Yaskawa INFORM job: VEGG1.JBI

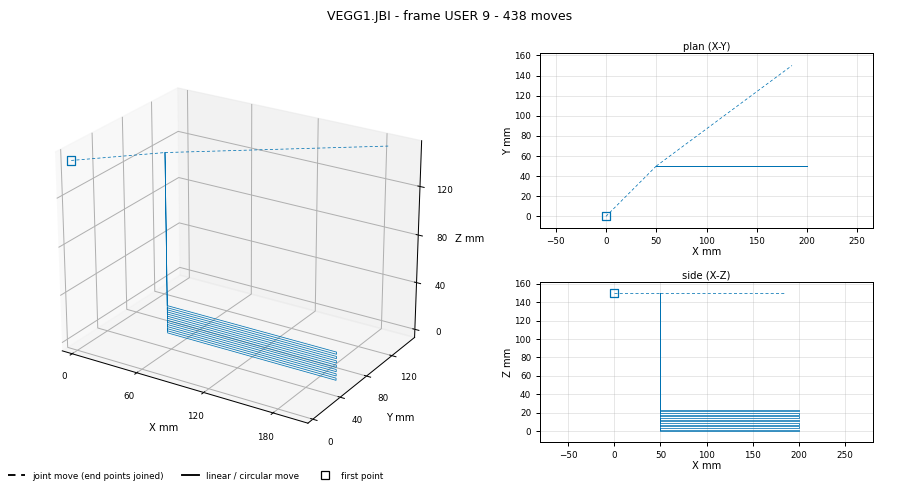
[picture p0: tool path of VEGG1.JBI in frame USER 9, 438 of 438 moves have a stored position in this frame; points joined in program order, loops and branches not executed]
/JOB
//NAME VEGG1
//POS
///NPOS 438,0,0,0,0,0
///USER 9
///TOOL 1
///POSTYPE USER
///RECTAN
///RCONF 1,0,0,0,0,0,0,0,0,0,0,0,0,0,0,0,0,0,0,0,0,0,0,0
C00000=0.000,0.000,150.000,0.0000,0.0000,180.0000
C00001=50.000,50.000,150.000,0.0000,0.0000,180.0000
C00002=50.000,50.000,0.000,0.0000,0.0000,180.0000
C00003=55.000,50.000,0.000,0.0000,0.0000,180.0000
C00004=60.000,50.000,0.000,0.0000,0.0000,180.0000
C00005=65.000,50.000,0.000,0.0000,0.0000,180.0000
C00006=70.000,50.000,0.000,0.0000,0.0000,180.0000
C00007=75.000,50.000,0.000,0.0000,0.0000,180.0000
C00008=80.000,50.000,0.000,0.0000,0.0000,180.0000
C00009=85.000,50.000,0.000,0.0000,0.0000,180.0000
C00010=90.000,50.000,0.000,0.0000,0.0000,180.0000
C00011=95.000,50.000,0.000,0.0000,0.0000,180.0000
C00012=100.000,50.000,0.000,0.0000,0.0000,180.0000
C00013=105.000,50.000,0.000,0.0000,0.0000,180.0000
C00014=110.000,50.000,0.000,0.0000,0.0000,180.0000
C00015=115.000,50.000,0.000,0.0000,0.0000,180.0000
C00016=120.000,50.000,0.000,0.0000,0.0000,180.0000
C00017=125.000,50.000,0.000,0.0000,0.0000,180.0000
C00018=130.000,50.000,0.000,0.0000,0.0000,180.0000
C00019=135.000,50.000,0.000,0.0000,0.0000,180.0000
C00020=140.000,50.000,0.000,0.0000,0.0000,180.0000
C00021=145.000,50.000,0.000,0.0000,0.0000,180.0000
C00022=150.000,50.000,0.000,0.0000,0.0000,180.0000
C00023=155.000,50.000,0.000,0.0000,0.0000,180.0000
C00024=160.000,50.000,0.000,0.0000,0.0000,180.0000
C00025=165.000,50.000,0.000,0.0000,0.0000,180.0000
C00026=170.000,50.000,0.000,0.0000,0.0000,180.0000
C00027=175.000,50.000,0.000,0.0000,0.0000,180.0000
C00028=180.000,50.000,0.000,0.0000,0.0000,180.0000
C00029=185.000,50.000,0.000,0.0000,0.0000,180.0000
C00030=190.000,50.000,0.000,0.0000,0.0000,180.0000
C00031=195.000,50.000,0.000,0.0000,0.0000,180.0000
C00032=200.000,50.000,0.000,0.0000,0.0000,180.0000
C00033=200.000,50.000,1.800,0.0000,0.0000,180.0000
C00034=195.000,50.000,1.800,0.0000,0.0000,180.0000
C00035=190.000,50.000,1.800,0.0000,0.0000,180.0000
C00036=185.000,50.000,1.800,0.0000,0.0000,180.0000
C00037=180.000,50.000,1.800,0.0000,0.0000,180.0000
C00038=175.000,50.000,1.800,0.0000,0.0000,180.0000
C00039=170.000,50.000,1.800,0.0000,0.0000,180.0000
C00040=165.000,50.000,1.800,0.0000,0.0000,180.0000
C00041=160.000,50.000,1.800,0.0000,0.0000,180.0000
C00042=155.000,50.000,1.800,0.0000,0.0000,180.0000
C00043=150.000,50.000,1.800,0.0000,0.0000,180.0000
C00044=145.000,50.000,1.800,0.0000,0.0000,180.0000
C00045=140.000,50.000,1.800,0.0000,0.0000,180.0000
C00046=135.000,50.000,1.800,0.0000,0.0000,180.0000
C00047=130.000,50.000,1.800,0.0000,0.0000,180.0000
C00048=125.000,50.000,1.800,0.0000,0.0000,180.0000
C00049=120.000,50.000,1.800,0.0000,0.0000,180.0000
C00050=115.000,50.000,1.800,0.0000,0.0000,180.0000
C00051=110.000,50.000,1.800,0.0000,0.0000,180.0000
C00052=105.000,50.000,1.800,0.0000,0.0000,180.0000
C00053=100.000,50.000,1.800,0.0000,0.0000,180.0000
C00054=95.000,50.000,1.800,0.0000,0.0000,180.0000
C00055=90.000,50.000,1.800,0.0000,0.0000,180.0000
C00056=85.000,50.000,1.800,0.0000,0.0000,180.0000
C00057=80.000,50.000,1.800,0.0000,0.0000,180.0000
C00058=75.000,50.000,1.800,0.0000,0.0000,180.0000
C00059=70.000,50.000,1.800,0.0000,0.0000,180.0000
C00060=65.000,50.000,1.800,0.0000,0.0000,180.0000
C00061=60.000,50.000,1.800,0.0000,0.0000,180.0000
C00062=55.000,50.000,1.800,0.0000,0.0000,180.0000
C00063=50.000,50.000,1.800,0.0000,0.0000,180.0000
C00064=50.000,50.000,3.600,0.0000,0.0000,180.0000
C00065=55.000,50.000,3.600,0.0000,0.0000,180.0000
C00066=60.000,50.000,3.600,0.0000,0.0000,180.0000
C00067=65.000,50.000,3.600,0.0000,0.0000,180.0000
C00068=70.000,50.000,3.600,0.0000,0.0000,180.0000
C00069=75.000,50.000,3.600,0.0000,0.0000,180.0000
C00070=80.000,50.000,3.600,0.0000,0.0000,180.0000
C00071=85.000,50.000,3.600,0.0000,0.0000,180.0000
C00072=90.000,50.000,3.600,0.0000,0.0000,180.0000
C00073=95.000,50.000,3.600,0.0000,0.0000,180.0000
C00074=100.000,50.000,3.600,0.0000,0.0000,180.0000
C00075=105.000,50.000,3.600,0.0000,0.0000,180.0000
C00076=110.000,50.000,3.600,0.0000,0.0000,180.0000
C00077=115.000,50.000,3.600,0.0000,0.0000,180.0000
C00078=120.000,50.000,3.600,0.0000,0.0000,180.0000
C00079=125.000,50.000,3.600,0.0000,0.0000,180.0000
C00080=130.000,50.000,3.600,0.0000,0.0000,180.0000
C00081=135.000,50.000,3.600,0.0000,0.0000,180.0000
C00082=140.000,50.000,3.600,0.0000,0.0000,180.0000
C00083=145.000,50.000,3.600,0.0000,0.0000,180.0000
C00084=150.000,50.000,3.600,0.0000,0.0000,180.0000
C00085=155.000,50.000,3.600,0.0000,0.0000,180.0000
C00086=160.000,50.000,3.600,0.0000,0.0000,180.0000
C00087=165.000,50.000,3.600,0.0000,0.0000,180.0000
C00088=170.000,50.000,3.600,0.0000,0.0000,180.0000
C00089=175.000,50.000,3.600,0.0000,0.0000,180.0000
C00090=180.000,50.000,3.600,0.0000,0.0000,180.0000
C00091=185.000,50.000,3.600,0.0000,0.0000,180.0000
C00092=190.000,50.000,3.600,0.0000,0.0000,180.0000
C00093=195.000,50.000,3.600,0.0000,0.0000,180.0000
C00094=200.000,50.000,3.600,0.0000,0.0000,180.0000
C00095=200.000,50.000,5.400,0.0000,0.0000,180.0000
C00096=195.000,50.000,5.400,0.0000,0.0000,180.0000
C00097=190.000,50.000,5.400,0.0000,0.0000,180.0000
C00098=185.000,50.000,5.400,0.0000,0.0000,180.0000
C00099=180.000,50.000,5.400,0.0000,0.0000,180.0000
C00100=175.000,50.000,5.400,0.0000,0.0000,180.0000
C00101=170.000,50.000,5.400,0.0000,0.0000,180.0000
C00102=165.000,50.000,5.400,0.0000,0.0000,180.0000
C00103=160.000,50.000,5.400,0.0000,0.0000,180.0000
C00104=155.000,50.000,5.400,0.0000,0.0000,180.0000
C00105=150.000,50.000,5.400,0.0000,0.0000,180.0000
C00106=145.000,50.000,5.400,0.0000,0.0000,180.0000
C00107=140.000,50.000,5.400,0.0000,0.0000,180.0000
C00108=135.000,50.000,5.400,0.0000,0.0000,180.0000
C00109=130.000,50.000,5.400,0.0000,0.0000,180.0000
C00110=125.000,50.000,5.400,0.0000,0.0000,180.0000
C00111=120.000,50.000,5.400,0.0000,0.0000,180.0000
C00112=115.000,50.000,5.400,0.0000,0.0000,180.0000
C00113=110.000,50.000,5.400,0.0000,0.0000,180.0000
C00114=105.000,50.000,5.400,0.0000,0.0000,180.0000
C00115=100.000,50.000,5.400,0.0000,0.0000,180.0000
C00116=95.000,50.000,5.400,0.0000,0.0000,180.0000
C00117=90.000,50.000,5.400,0.0000,0.0000,180.0000
C00118=85.000,50.000,5.400,0.0000,0.0000,180.0000
C00119=80.000,50.000,5.400,0.0000,0.0000,180.0000
C00120=75.000,50.000,5.400,0.0000,0.0000,180.0000
C00121=70.000,50.000,5.400,0.0000,0.0000,180.0000
C00122=65.000,50.000,5.400,0.0000,0.0000,180.0000
C00123=60.000,50.000,5.400,0.0000,0.0000,180.0000
C00124=55.000,50.000,5.400,0.0000,0.0000,180.0000
C00125=50.000,50.000,5.400,0.0000,0.0000,180.0000
C00126=50.000,50.000,7.200,0.0000,0.0000,180.0000
C00127=55.000,50.000,7.200,0.0000,0.0000,180.0000
C00128=60.000,50.000,7.200,0.0000,0.0000,180.0000
C00129=65.000,50.000,7.200,0.0000,0.0000,180.0000
C00130=70.000,50.000,7.200,0.0000,0.0000,180.0000
C00131=75.000,50.000,7.200,0.0000,0.0000,180.0000
C00132=80.000,50.000,7.200,0.0000,0.0000,180.0000
C00133=85.000,50.000,7.200,0.0000,0.0000,180.0000
C00134=90.000,50.000,7.200,0.0000,0.0000,180.0000
C00135=95.000,50.000,7.200,0.0000,0.0000,180.0000
C00136=100.000,50.000,7.200,0.0000,0.0000,180.0000
C00137=105.000,50.000,7.200,0.0000,0.0000,180.0000
C00138=110.000,50.000,7.200,0.0000,0.0000,180.0000
C00139=115.000,50.000,7.200,0.0000,0.0000,180.0000
C00140=120.000,50.000,7.200,0.0000,0.0000,180.0000
C00141=125.000,50.000,7.200,0.0000,0.0000,180.0000
C00142=130.000,50.000,7.200,0.0000,0.0000,180.0000
C00143=135.000,50.000,7.200,0.0000,0.0000,180.0000
C00144=140.000,50.000,7.200,0.0000,0.0000,180.0000
C00145=145.000,50.000,7.200,0.0000,0.0000,180.0000
C00146=150.000,50.000,7.200,0.0000,0.0000,180.0000
C00147=155.000,50.000,7.200,0.0000,0.0000,180.0000
C00148=160.000,50.000,7.200,0.0000,0.0000,180.0000
C00149=165.000,50.000,7.200,0.0000,0.0000,180.0000
C00150=170.000,50.000,7.200,0.0000,0.0000,180.0000
C00151=175.000,50.000,7.200,0.0000,0.0000,180.0000
C00152=180.000,50.000,7.200,0.0000,0.0000,180.0000
C00153=185.000,50.000,7.200,0.0000,0.0000,180.0000
C00154=190.000,50.000,7.200,0.0000,0.0000,180.0000
C00155=195.000,50.000,7.200,0.0000,0.0000,180.0000
C00156=200.000,50.000,7.200,0.0000,0.0000,180.0000
C00157=200.000,50.000,9.000,0.0000,0.0000,180.0000
C00158=195.000,50.000,9.000,0.0000,0.0000,180.0000
C00159=190.000,50.000,9.000,0.0000,0.0000,180.0000
C00160=185.000,50.000,9.000,0.0000,0.0000,180.0000
C00161=180.000,50.000,9.000,0.0000,0.0000,180.0000
C00162=175.000,50.000,9.000,0.0000,0.0000,180.0000
C00163=170.000,50.000,9.000,0.0000,0.0000,180.0000
C00164=165.000,50.000,9.000,0.0000,0.0000,180.0000
C00165=160.000,50.000,9.000,0.0000,0.0000,180.0000
C00166=155.000,50.000,9.000,0.0000,0.0000,180.0000
C00167=150.000,50.000,9.000,0.0000,0.0000,180.0000
C00168=145.000,50.000,9.000,0.0000,0.0000,180.0000
C00169=140.000,50.000,9.000,0.0000,0.0000,180.0000
C00170=135.000,50.000,9.000,0.0000,0.0000,180.0000
C00171=130.000,50.000,9.000,0.0000,0.0000,180.0000
C00172=125.000,50.000,9.000,0.0000,0.0000,180.0000
C00173=120.000,50.000,9.000,0.0000,0.0000,180.0000
C00174=115.000,50.000,9.000,0.0000,0.0000,180.0000
C00175=110.000,50.000,9.000,0.0000,0.0000,180.0000
C00176=105.000,50.000,9.000,0.0000,0.0000,180.0000
C00177=100.000,50.000,9.000,0.0000,0.0000,180.0000
C00178=95.000,50.000,9.000,0.0000,0.0000,180.0000
C00179=90.000,50.000,9.000,0.0000,0.0000,180.0000
C00180=85.000,50.000,9.000,0.0000,0.0000,180.0000
C00181=80.000,50.000,9.000,0.0000,0.0000,180.0000
C00182=75.000,50.000,9.000,0.0000,0.0000,180.0000
C00183=70.000,50.000,9.000,0.0000,0.0000,180.0000
C00184=65.000,50.000,9.000,0.0000,0.0000,180.0000
C00185=60.000,50.000,9.000,0.0000,0.0000,180.0000
C00186=55.000,50.000,9.000,0.0000,0.0000,180.0000
C00187=50.000,50.000,9.000,0.0000,0.0000,180.0000
C00188=50.000,50.000,10.800,0.0000,0.0000,180.0000
C00189=55.000,50.000,10.800,0.0000,0.0000,180.0000
C00190=60.000,50.000,10.800,0.0000,0.0000,180.0000
C00191=65.000,50.000,10.800,0.0000,0.0000,180.0000
C00192=70.000,50.000,10.800,0.0000,0.0000,180.0000
C00193=75.000,50.000,10.800,0.0000,0.0000,180.0000
C00194=80.000,50.000,10.800,0.0000,0.0000,180.0000
C00195=85.000,50.000,10.800,0.0000,0.0000,180.0000
C00196=90.000,50.000,10.800,0.0000,0.0000,180.0000
C00197=95.000,50.000,10.800,0.0000,0.0000,180.0000
C00198=100.000,50.000,10.800,0.0000,0.0000,180.0000
C00199=105.000,50.000,10.800,0.0000,0.0000,180.0000
C00200=110.000,50.000,10.800,0.0000,0.0000,180.0000
C00201=115.000,50.000,10.800,0.0000,0.0000,180.0000
C00202=120.000,50.000,10.800,0.0000,0.0000,180.0000
C00203=125.000,50.000,10.800,0.0000,0.0000,180.0000
C00204=130.000,50.000,10.800,0.0000,0.0000,180.0000
C00205=135.000,50.000,10.800,0.0000,0.0000,180.0000
C00206=140.000,50.000,10.800,0.0000,0.0000,180.0000
C00207=145.000,50.000,10.800,0.0000,0.0000,180.0000
C00208=150.000,50.000,10.800,0.0000,0.0000,180.0000
C00209=155.000,50.000,10.800,0.0000,0.0000,180.0000
C00210=160.000,50.000,10.800,0.0000,0.0000,180.0000
C00211=165.000,50.000,10.800,0.0000,0.0000,180.0000
C00212=170.000,50.000,10.800,0.0000,0.0000,180.0000
C00213=175.000,50.000,10.800,0.0000,0.0000,180.0000
C00214=180.000,50.000,10.800,0.0000,0.0000,180.0000
C00215=185.000,50.000,10.800,0.0000,0.0000,180.0000
C00216=190.000,50.000,10.800,0.0000,0.0000,180.0000
C00217=195.000,50.000,10.800,0.0000,0.0000,180.0000
C00218=200.000,50.000,10.800,0.0000,0.0000,180.0000
C00219=200.000,50.000,12.600,0.0000,0.0000,180.0000
C00220=195.000,50.000,12.600,0.0000,0.0000,180.0000
C00221=190.000,50.000,12.600,0.0000,0.0000,180.0000
C00222=185.000,50.000,12.600,0.0000,0.0000,180.0000
C00223=180.000,50.000,12.600,0.0000,0.0000,180.0000
C00224=175.000,50.000,12.600,0.0000,0.0000,180.0000
C00225=170.000,50.000,12.600,0.0000,0.0000,180.0000
C00226=165.000,50.000,12.600,0.0000,0.0000,180.0000
C00227=160.000,50.000,12.600,0.0000,0.0000,180.0000
C00228=155.000,50.000,12.600,0.0000,0.0000,180.0000
C00229=150.000,50.000,12.600,0.0000,0.0000,180.0000
C00230=145.000,50.000,12.600,0.0000,0.0000,180.0000
C00231=140.000,50.000,12.600,0.0000,0.0000,180.0000
C00232=135.000,50.000,12.600,0.0000,0.0000,180.0000
C00233=130.000,50.000,12.600,0.0000,0.0000,180.0000
C00234=125.000,50.000,12.600,0.0000,0.0000,180.0000
C00235=120.000,50.000,12.600,0.0000,0.0000,180.0000
C00236=115.000,50.000,12.600,0.0000,0.0000,180.0000
C00237=110.000,50.000,12.600,0.0000,0.0000,180.0000
C00238=105.000,50.000,12.600,0.0000,0.0000,180.0000
C00239=100.000,50.000,12.600,0.0000,0.0000,180.0000
C00240=95.000,50.000,12.600,0.0000,0.0000,180.0000
C00241=90.000,50.000,12.600,0.0000,0.0000,180.0000
C00242=85.000,50.000,12.600,0.0000,0.0000,180.0000
C00243=80.000,50.000,12.600,0.0000,0.0000,180.0000
C00244=75.000,50.000,12.600,0.0000,0.0000,180.0000
C00245=70.000,50.000,12.600,0.0000,0.0000,180.0000
C00246=65.000,50.000,12.600,0.0000,0.0000,180.0000
C00247=60.000,50.000,12.600,0.0000,0.0000,180.0000
C00248=55.000,50.000,12.600,0.0000,0.0000,180.0000
C00249=50.000,50.000,12.600,0.0000,0.0000,180.0000
C00250=50.000,50.000,14.400,0.0000,0.0000,180.0000
C00251=55.000,50.000,14.400,0.0000,0.0000,180.0000
C00252=60.000,50.000,14.400,0.0000,0.0000,180.0000
C00253=65.000,50.000,14.400,0.0000,0.0000,180.0000
C00254=70.000,50.000,14.400,0.0000,0.0000,180.0000
C00255=75.000,50.000,14.400,0.0000,0.0000,180.0000
C00256=80.000,50.000,14.400,0.0000,0.0000,180.0000
C00257=85.000,50.000,14.400,0.0000,0.0000,180.0000
C00258=90.000,50.000,14.400,0.0000,0.0000,180.0000
C00259=95.000,50.000,14.400,0.0000,0.0000,180.0000
C00260=100.000,50.000,14.400,0.0000,0.0000,180.0000
C00261=105.000,50.000,14.400,0.0000,0.0000,180.0000
C00262=110.000,50.000,14.400,0.0000,0.0000,180.0000
C00263=115.000,50.000,14.400,0.0000,0.0000,180.0000
C00264=120.000,50.000,14.400,0.0000,0.0000,180.0000
C00265=125.000,50.000,14.400,0.0000,0.0000,180.0000
C00266=130.000,50.000,14.400,0.0000,0.0000,180.0000
C00267=135.000,50.000,14.400,0.0000,0.0000,180.0000
C00268=140.000,50.000,14.400,0.0000,0.0000,180.0000
C00269=145.000,50.000,14.400,0.0000,0.0000,180.0000
C00270=150.000,50.000,14.400,0.0000,0.0000,180.0000
C00271=155.000,50.000,14.400,0.0000,0.0000,180.0000
C00272=160.000,50.000,14.400,0.0000,0.0000,180.0000
C00273=165.000,50.000,14.400,0.0000,0.0000,180.0000
C00274=170.000,50.000,14.400,0.0000,0.0000,180.0000
C00275=175.000,50.000,14.400,0.0000,0.0000,180.0000
C00276=180.000,50.000,14.400,0.0000,0.0000,180.0000
C00277=185.000,50.000,14.400,0.0000,0.0000,180.0000
C00278=190.000,50.000,14.400,0.0000,0.0000,180.0000
C00279=195.000,50.000,14.400,0.0000,0.0000,180.0000
C00280=200.000,50.000,14.400,0.0000,0.0000,180.0000
C00281=200.000,50.000,16.200,0.0000,0.0000,180.0000
C00282=195.000,50.000,16.200,0.0000,0.0000,180.0000
C00283=190.000,50.000,16.200,0.0000,0.0000,180.0000
C00284=185.000,50.000,16.200,0.0000,0.0000,180.0000
C00285=180.000,50.000,16.200,0.0000,0.0000,180.0000
C00286=175.000,50.000,16.200,0.0000,0.0000,180.0000
C00287=170.000,50.000,16.200,0.0000,0.0000,180.0000
C00288=165.000,50.000,16.200,0.0000,0.0000,180.0000
C00289=160.000,50.000,16.200,0.0000,0.0000,180.0000
C00290=155.000,50.000,16.200,0.0000,0.0000,180.0000
C00291=150.000,50.000,16.200,0.0000,0.0000,180.0000
C00292=145.000,50.000,16.200,0.0000,0.0000,180.0000
C00293=140.000,50.000,16.200,0.0000,0.0000,180.0000
C00294=135.000,50.000,16.200,0.0000,0.0000,180.0000
C00295=130.000,50.000,16.200,0.0000,0.0000,180.0000
C00296=125.000,50.000,16.200,0.0000,0.0000,180.0000
C00297=120.000,50.000,16.200,0.0000,0.0000,180.0000
C00298=115.000,50.000,16.200,0.0000,0.0000,180.0000
C00299=110.000,50.000,16.200,0.0000,0.0000,180.0000
C00300=105.000,50.000,16.200,0.0000,0.0000,180.0000
C00301=100.000,50.000,16.200,0.0000,0.0000,180.0000
C00302=95.000,50.000,16.200,0.0000,0.0000,180.0000
C00303=90.000,50.000,16.200,0.0000,0.0000,180.0000
C00304=85.000,50.000,16.200,0.0000,0.0000,180.0000
C00305=80.000,50.000,16.200,0.0000,0.0000,180.0000
C00306=75.000,50.000,16.200,0.0000,0.0000,180.0000
C00307=70.000,50.000,16.200,0.0000,0.0000,180.0000
C00308=65.000,50.000,16.200,0.0000,0.0000,180.0000
C00309=60.000,50.000,16.200,0.0000,0.0000,180.0000
C00310=55.000,50.000,16.200,0.0000,0.0000,180.0000
C00311=50.000,50.000,16.200,0.0000,0.0000,180.0000
C00312=50.000,50.000,18.000,0.0000,0.0000,180.0000
C00313=55.000,50.000,18.000,0.0000,0.0000,180.0000
C00314=60.000,50.000,18.000,0.0000,0.0000,180.0000
C00315=65.000,50.000,18.000,0.0000,0.0000,180.0000
C00316=70.000,50.000,18.000,0.0000,0.0000,180.0000
C00317=75.000,50.000,18.000,0.0000,0.0000,180.0000
C00318=80.000,50.000,18.000,0.0000,0.0000,180.0000
C00319=85.000,50.000,18.000,0.0000,0.0000,180.0000
C00320=90.000,50.000,18.000,0.0000,0.0000,180.0000
C00321=95.000,50.000,18.000,0.0000,0.0000,180.0000
C00322=100.000,50.000,18.000,0.0000,0.0000,180.0000
C00323=105.000,50.000,18.000,0.0000,0.0000,180.0000
C00324=110.000,50.000,18.000,0.0000,0.0000,180.0000
C00325=115.000,50.000,18.000,0.0000,0.0000,180.0000
C00326=120.000,50.000,18.000,0.0000,0.0000,180.0000
C00327=125.000,50.000,18.000,0.0000,0.0000,180.0000
C00328=130.000,50.000,18.000,0.0000,0.0000,180.0000
C00329=135.000,50.000,18.000,0.0000,0.0000,180.0000
C00330=140.000,50.000,18.000,0.0000,0.0000,180.0000
C00331=145.000,50.000,18.000,0.0000,0.0000,180.0000
C00332=150.000,50.000,18.000,0.0000,0.0000,180.0000
C00333=155.000,50.000,18.000,0.0000,0.0000,180.0000
C00334=160.000,50.000,18.000,0.0000,0.0000,180.0000
C00335=165.000,50.000,18.000,0.0000,0.0000,180.0000
C00336=170.000,50.000,18.000,0.0000,0.0000,180.0000
C00337=175.000,50.000,18.000,0.0000,0.0000,180.0000
C00338=180.000,50.000,18.000,0.0000,0.0000,180.0000
C00339=185.000,50.000,18.000,0.0000,0.0000,180.0000
C00340=190.000,50.000,18.000,0.0000,0.0000,180.0000
C00341=195.000,50.000,18.000,0.0000,0.0000,180.0000
C00342=200.000,50.000,18.000,0.0000,0.0000,180.0000
C00343=200.000,50.000,19.800,0.0000,0.0000,180.0000
C00344=195.000,50.000,19.800,0.0000,0.0000,180.0000
C00345=190.000,50.000,19.800,0.0000,0.0000,180.0000
C00346=185.000,50.000,19.800,0.0000,0.0000,180.0000
C00347=180.000,50.000,19.800,0.0000,0.0000,180.0000
C00348=175.000,50.000,19.800,0.0000,0.0000,180.0000
C00349=170.000,50.000,19.800,0.0000,0.0000,180.0000
C00350=165.000,50.000,19.800,0.0000,0.0000,180.0000
C00351=160.000,50.000,19.800,0.0000,0.0000,180.0000
C00352=155.000,50.000,19.800,0.0000,0.0000,180.0000
C00353=150.000,50.000,19.800,0.0000,0.0000,180.0000
C00354=145.000,50.000,19.800,0.0000,0.0000,180.0000
C00355=140.000,50.000,19.800,0.0000,0.0000,180.0000
C00356=135.000,50.000,19.800,0.0000,0.0000,180.0000
C00357=130.000,50.000,19.800,0.0000,0.0000,180.0000
C00358=125.000,50.000,19.800,0.0000,0.0000,180.0000
C00359=120.000,50.000,19.800,0.0000,0.0000,180.0000
C00360=115.000,50.000,19.800,0.0000,0.0000,180.0000
C00361=110.000,50.000,19.800,0.0000,0.0000,180.0000
C00362=105.000,50.000,19.800,0.0000,0.0000,180.0000
C00363=100.000,50.000,19.800,0.0000,0.0000,180.0000
C00364=95.000,50.000,19.800,0.0000,0.0000,180.0000
C00365=90.000,50.000,19.800,0.0000,0.0000,180.0000
C00366=85.000,50.000,19.800,0.0000,0.0000,180.0000
C00367=80.000,50.000,19.800,0.0000,0.0000,180.0000
C00368=75.000,50.000,19.800,0.0000,0.0000,180.0000
C00369=70.000,50.000,19.800,0.0000,0.0000,180.0000
C00370=65.000,50.000,19.800,0.0000,0.0000,180.0000
C00371=60.000,50.000,19.800,0.0000,0.0000,180.0000
C00372=55.000,50.000,19.800,0.0000,0.0000,180.0000
C00373=50.000,50.000,19.800,0.0000,0.0000,180.0000
C00374=50.000,50.000,21.600,0.0000,0.0000,180.0000
C00375=55.000,50.000,21.600,0.0000,0.0000,180.0000
C00376=60.000,50.000,21.600,0.0000,0.0000,180.0000
C00377=65.000,50.000,21.600,0.0000,0.0000,180.0000
C00378=70.000,50.000,21.600,0.0000,0.0000,180.0000
C00379=75.000,50.000,21.600,0.0000,0.0000,180.0000
C00380=80.000,50.000,21.600,0.0000,0.0000,180.0000
C00381=85.000,50.000,21.600,0.0000,0.0000,180.0000
C00382=90.000,50.000,21.600,0.0000,0.0000,180.0000
C00383=95.000,50.000,21.600,0.0000,0.0000,180.0000
C00384=100.000,50.000,21.600,0.0000,0.0000,180.0000
C00385=105.000,50.000,21.600,0.0000,0.0000,180.0000
C00386=110.000,50.000,21.600,0.0000,0.0000,180.0000
C00387=115.000,50.000,21.600,0.0000,0.0000,180.0000
C00388=120.000,50.000,21.600,0.0000,0.0000,180.0000
C00389=125.000,50.000,21.600,0.0000,0.0000,180.0000
C00390=130.000,50.000,21.600,0.0000,0.0000,180.0000
C00391=135.000,50.000,21.600,0.0000,0.0000,180.0000
C00392=140.000,50.000,21.600,0.0000,0.0000,180.0000
C00393=145.000,50.000,21.600,0.0000,0.0000,180.0000
C00394=150.000,50.000,21.600,0.0000,0.0000,180.0000
C00395=155.000,50.000,21.600,0.0000,0.0000,180.0000
C00396=160.000,50.000,21.600,0.0000,0.0000,180.0000
C00397=165.000,50.000,21.600,0.0000,0.0000,180.0000
C00398=170.000,50.000,21.600,0.0000,0.0000,180.0000
C00399=175.000,50.000,21.600,0.0000,0.0000,180.0000
C00400=180.000,50.000,21.600,0.0000,0.0000,180.0000
C00401=185.000,50.000,21.600,0.0000,0.0000,180.0000
C00402=190.000,50.000,21.600,0.0000,0.0000,180.0000
C00403=195.000,50.000,21.600,0.0000,0.0000,180.0000
C00404=200.000,50.000,21.600,0.0000,0.0000,180.0000
C00405=200.000,50.000,23.400,0.0000,0.0000,180.0000
C00406=195.000,50.000,23.400,0.0000,0.0000,180.0000
C00407=190.000,50.000,23.400,0.0000,0.0000,180.0000
C00408=185.000,50.000,23.400,0.0000,0.0000,180.0000
C00409=180.000,50.000,23.400,0.0000,0.0000,180.0000
C00410=175.000,50.000,23.400,0.0000,0.0000,180.0000
C00411=170.000,50.000,23.400,0.0000,0.0000,180.0000
C00412=165.000,50.000,23.400,0.0000,0.0000,180.0000
C00413=160.000,50.000,23.400,0.0000,0.0000,180.0000
C00414=155.000,50.000,23.400,0.0000,0.0000,180.0000
C00415=150.000,50.000,23.400,0.0000,0.0000,180.0000
C00416=145.000,50.000,23.400,0.0000,0.0000,180.0000
C00417=140.000,50.000,23.400,0.0000,0.0000,180.0000
C00418=135.000,50.000,23.400,0.0000,0.0000,180.0000
C00419=130.000,50.000,23.400,0.0000,0.0000,180.0000
C00420=125.000,50.000,23.400,0.0000,0.0000,180.0000
C00421=120.000,50.000,23.400,0.0000,0.0000,180.0000
C00422=115.000,50.000,23.400,0.0000,0.0000,180.0000
C00423=110.000,50.000,23.400,0.0000,0.0000,180.0000
C00424=105.000,50.000,23.400,0.0000,0.0000,180.0000
C00425=100.000,50.000,23.400,0.0000,0.0000,180.0000
C00426=95.000,50.000,23.400,0.0000,0.0000,180.0000
C00427=90.000,50.000,23.400,0.0000,0.0000,180.0000
C00428=85.000,50.000,23.400,0.0000,0.0000,180.0000
C00429=80.000,50.000,23.400,0.0000,0.0000,180.0000
C00430=75.000,50.000,23.400,0.0000,0.0000,180.0000
C00431=70.000,50.000,23.400,0.0000,0.0000,180.0000
C00432=65.000,50.000,23.400,0.0000,0.0000,180.0000
C00433=60.000,50.000,23.400,0.0000,0.0000,180.0000
C00434=55.000,50.000,23.400,0.0000,0.0000,180.0000
C00435=50.000,50.000,23.400,0.0000,0.0000,180.0000
C00436=50.000,50.000,150.000,0.0000,0.0000,180.0000
C00437=185.000,150.000,150.000,0.0000,0.0000,180.0000
//INST
///DATE 2026/10/20 11:28
///ATTR SC,RW,RJ
////FRAME USER 9
///GROUP1 RB1
NOP
MOVJ C00000 VJ=0.78
MOVJ C00001 VJ=0.78
MOVL C00002 V=11.0 ACC=20 DEC=20
MACRO1 MJ#(0) ARGF1
ARCON
MOVL C00003 V=8.0 ACC=20 DEC=20
MOVL C00004 V=8.0 ACC=20 DEC=20
MOVL C00005 V=8.0 ACC=20 DEC=20
MOVL C00006 V=8.0 ACC=20 DEC=20
MOVL C00007 V=8.0 ACC=20 DEC=20
MOVL C00008 V=8.0 ACC=20 DEC=20
MOVL C00009 V=8.0 ACC=20 DEC=20
MOVL C00010 V=8.0 ACC=20 DEC=20
MOVL C00011 V=8.0 ACC=20 DEC=20
MOVL C00012 V=8.0 ACC=20 DEC=20
MOVL C00013 V=8.0 ACC=20 DEC=20
MOVL C00014 V=8.0 ACC=20 DEC=20
MOVL C00015 V=8.0 ACC=20 DEC=20
MOVL C00016 V=8.0 ACC=20 DEC=20
MOVL C00017 V=8.0 ACC=20 DEC=20
MOVL C00018 V=8.0 ACC=20 DEC=20
MOVL C00019 V=8.0 ACC=20 DEC=20
MOVL C00020 V=8.0 ACC=20 DEC=20
MOVL C00021 V=8.0 ACC=20 DEC=20
MOVL C00022 V=8.0 ACC=20 DEC=20
MOVL C00023 V=8.0 ACC=20 DEC=20
MOVL C00024 V=8.0 ACC=20 DEC=20
MOVL C00025 V=8.0 ACC=20 DEC=20
MOVL C00026 V=8.0 ACC=20 DEC=20
MOVL C00027 V=8.0 ACC=20 DEC=20
MOVL C00028 V=8.0 ACC=20 DEC=20
MOVL C00029 V=8.0 ACC=20 DEC=20
MOVL C00030 V=8.0 ACC=20 DEC=20
MOVL C00031 V=8.0 ACC=20 DEC=20
MOVL C00032 V=8.0 ACC=20 DEC=20
ARCOF
TIMER T=60.0
MOVL C00033 V=11.0 ACC=20 DEC=20
MACRO1 MJ#(0) ARGF2
ARCON
MOVL C00034 V=8.0 ACC=20 DEC=20
MOVL C00035 V=8.0 ACC=20 DEC=20
MOVL C00036 V=8.0 ACC=20 DEC=20
MOVL C00037 V=8.0 ACC=20 DEC=20
MOVL C00038 V=8.0 ACC=20 DEC=20
MOVL C00039 V=8.0 ACC=20 DEC=20
MOVL C00040 V=8.0 ACC=20 DEC=20
MOVL C00041 V=8.0 ACC=20 DEC=20
MOVL C00042 V=8.0 ACC=20 DEC=20
MOVL C00043 V=8.0 ACC=20 DEC=20
MOVL C00044 V=8.0 ACC=20 DEC=20
MOVL C00045 V=8.0 ACC=20 DEC=20
MOVL C00046 V=8.0 ACC=20 DEC=20
MOVL C00047 V=8.0 ACC=20 DEC=20
MOVL C00048 V=8.0 ACC=20 DEC=20
MOVL C00049 V=8.0 ACC=20 DEC=20
MOVL C00050 V=8.0 ACC=20 DEC=20
MOVL C00051 V=8.0 ACC=20 DEC=20
MOVL C00052 V=8.0 ACC=20 DEC=20
MOVL C00053 V=8.0 ACC=20 DEC=20
MOVL C00054 V=8.0 ACC=20 DEC=20
MOVL C00055 V=8.0 ACC=20 DEC=20
MOVL C00056 V=8.0 ACC=20 DEC=20
MOVL C00057 V=8.0 ACC=20 DEC=20
MOVL C00058 V=8.0 ACC=20 DEC=20
MOVL C00059 V=8.0 ACC=20 DEC=20
MOVL C00060 V=8.0 ACC=20 DEC=20
MOVL C00061 V=8.0 ACC=20 DEC=20
MOVL C00062 V=8.0 ACC=20 DEC=20
MOVL C00063 V=8.0 ACC=20 DEC=20
ARCOF
TIMER T=60.0
MOVL C00064 V=11.0 ACC=20 DEC=20
MACRO1 MJ#(0) ARGF2
ARCON
MOVL C00065 V=8.0 ACC=20 DEC=20
MOVL C00066 V=8.0 ACC=20 DEC=20
MOVL C00067 V=8.0 ACC=20 DEC=20
MOVL C00068 V=8.0 ACC=20 DEC=20
MOVL C00069 V=8.0 ACC=20 DEC=20
MOVL C00070 V=8.0 ACC=20 DEC=20
MOVL C00071 V=8.0 ACC=20 DEC=20
MOVL C00072 V=8.0 ACC=20 DEC=20
MOVL C00073 V=8.0 ACC=20 DEC=20
MOVL C00074 V=8.0 ACC=20 DEC=20
MOVL C00075 V=8.0 ACC=20 DEC=20
MOVL C00076 V=8.0 ACC=20 DEC=20
MOVL C00077 V=8.0 ACC=20 DEC=20
MOVL C00078 V=8.0 ACC=20 DEC=20
MOVL C00079 V=8.0 ACC=20 DEC=20
MOVL C00080 V=8.0 ACC=20 DEC=20
MOVL C00081 V=8.0 ACC=20 DEC=20
MOVL C00082 V=8.0 ACC=20 DEC=20
MOVL C00083 V=8.0 ACC=20 DEC=20
MOVL C00084 V=8.0 ACC=20 DEC=20
MOVL C00085 V=8.0 ACC=20 DEC=20
MOVL C00086 V=8.0 ACC=20 DEC=20
MOVL C00087 V=8.0 ACC=20 DEC=20
MOVL C00088 V=8.0 ACC=20 DEC=20
MOVL C00089 V=8.0 ACC=20 DEC=20
MOVL C00090 V=8.0 ACC=20 DEC=20
MOVL C00091 V=8.0 ACC=20 DEC=20
MOVL C00092 V=8.0 ACC=20 DEC=20
MOVL C00093 V=8.0 ACC=20 DEC=20
MOVL C00094 V=8.0 ACC=20 DEC=20
ARCOF
TIMER T=60.0
MOVL C00095 V=11.0 ACC=20 DEC=20
MACRO1 MJ#(0) ARGF2
ARCON
MOVL C00096 V=8.0 ACC=20 DEC=20
MOVL C00097 V=8.0 ACC=20 DEC=20
MOVL C00098 V=8.0 ACC=20 DEC=20
MOVL C00099 V=8.0 ACC=20 DEC=20
MOVL C00100 V=8.0 ACC=20 DEC=20
MOVL C00101 V=8.0 ACC=20 DEC=20
MOVL C00102 V=8.0 ACC=20 DEC=20
MOVL C00103 V=8.0 ACC=20 DEC=20
MOVL C00104 V=8.0 ACC=20 DEC=20
MOVL C00105 V=8.0 ACC=20 DEC=20
MOVL C00106 V=8.0 ACC=20 DEC=20
MOVL C00107 V=8.0 ACC=20 DEC=20
MOVL C00108 V=8.0 ACC=20 DEC=20
MOVL C00109 V=8.0 ACC=20 DEC=20
MOVL C00110 V=8.0 ACC=20 DEC=20
MOVL C00111 V=8.0 ACC=20 DEC=20
MOVL C00112 V=8.0 ACC=20 DEC=20
MOVL C00113 V=8.0 ACC=20 DEC=20
MOVL C00114 V=8.0 ACC=20 DEC=20
MOVL C00115 V=8.0 ACC=20 DEC=20
MOVL C00116 V=8.0 ACC=20 DEC=20
MOVL C00117 V=8.0 ACC=20 DEC=20
MOVL C00118 V=8.0 ACC=20 DEC=20
MOVL C00119 V=8.0 ACC=20 DEC=20
MOVL C00120 V=8.0 ACC=20 DEC=20
MOVL C00121 V=8.0 ACC=20 DEC=20
MOVL C00122 V=8.0 ACC=20 DEC=20
MOVL C00123 V=8.0 ACC=20 DEC=20
MOVL C00124 V=8.0 ACC=20 DEC=20
MOVL C00125 V=8.0 ACC=20 DEC=20
ARCOF
TIMER T=60.0
MOVL C00126 V=11.0 ACC=20 DEC=20
MACRO1 MJ#(0) ARGF2
ARCON
MOVL C00127 V=8.0 ACC=20 DEC=20
MOVL C00128 V=8.0 ACC=20 DEC=20
MOVL C00129 V=8.0 ACC=20 DEC=20
MOVL C00130 V=8.0 ACC=20 DEC=20
MOVL C00131 V=8.0 ACC=20 DEC=20
MOVL C00132 V=8.0 ACC=20 DEC=20
MOVL C00133 V=8.0 ACC=20 DEC=20
MOVL C00134 V=8.0 ACC=20 DEC=20
MOVL C00135 V=8.0 ACC=20 DEC=20
MOVL C00136 V=8.0 ACC=20 DEC=20
MOVL C00137 V=8.0 ACC=20 DEC=20
MOVL C00138 V=8.0 ACC=20 DEC=20
MOVL C00139 V=8.0 ACC=20 DEC=20
MOVL C00140 V=8.0 ACC=20 DEC=20
MOVL C00141 V=8.0 ACC=20 DEC=20
MOVL C00142 V=8.0 ACC=20 DEC=20
MOVL C00143 V=8.0 ACC=20 DEC=20
MOVL C00144 V=8.0 ACC=20 DEC=20
MOVL C00145 V=8.0 ACC=20 DEC=20
MOVL C00146 V=8.0 ACC=20 DEC=20
MOVL C00147 V=8.0 ACC=20 DEC=20
MOVL C00148 V=8.0 ACC=20 DEC=20
MOVL C00149 V=8.0 ACC=20 DEC=20
MOVL C00150 V=8.0 ACC=20 DEC=20
MOVL C00151 V=8.0 ACC=20 DEC=20
MOVL C00152 V=8.0 ACC=20 DEC=20
MOVL C00153 V=8.0 ACC=20 DEC=20
MOVL C00154 V=8.0 ACC=20 DEC=20
MOVL C00155 V=8.0 ACC=20 DEC=20
MOVL C00156 V=8.0 ACC=20 DEC=20
ARCOF
TIMER T=60.0
MOVL C00157 V=11.0 ACC=20 DEC=20
MACRO1 MJ#(0) ARGF2
ARCON
MOVL C00158 V=8.0 ACC=20 DEC=20
MOVL C00159 V=8.0 ACC=20 DEC=20
MOVL C00160 V=8.0 ACC=20 DEC=20
MOVL C00161 V=8.0 ACC=20 DEC=20
MOVL C00162 V=8.0 ACC=20 DEC=20
MOVL C00163 V=8.0 ACC=20 DEC=20
MOVL C00164 V=8.0 ACC=20 DEC=20
MOVL C00165 V=8.0 ACC=20 DEC=20
MOVL C00166 V=8.0 ACC=20 DEC=20
MOVL C00167 V=8.0 ACC=20 DEC=20
MOVL C00168 V=8.0 ACC=20 DEC=20
MOVL C00169 V=8.0 ACC=20 DEC=20
MOVL C00170 V=8.0 ACC=20 DEC=20
MOVL C00171 V=8.0 ACC=20 DEC=20
MOVL C00172 V=8.0 ACC=20 DEC=20
MOVL C00173 V=8.0 ACC=20 DEC=20
MOVL C00174 V=8.0 ACC=20 DEC=20
MOVL C00175 V=8.0 ACC=20 DEC=20
MOVL C00176 V=8.0 ACC=20 DEC=20
MOVL C00177 V=8.0 ACC=20 DEC=20
MOVL C00178 V=8.0 ACC=20 DEC=20
MOVL C00179 V=8.0 ACC=20 DEC=20
MOVL C00180 V=8.0 ACC=20 DEC=20
MOVL C00181 V=8.0 ACC=20 DEC=20
MOVL C00182 V=8.0 ACC=20 DEC=20
MOVL C00183 V=8.0 ACC=20 DEC=20
MOVL C00184 V=8.0 ACC=20 DEC=20
MOVL C00185 V=8.0 ACC=20 DEC=20
MOVL C00186 V=8.0 ACC=20 DEC=20
MOVL C00187 V=8.0 ACC=20 DEC=20
ARCOF
TIMER T=60.0
MOVL C00188 V=11.0 ACC=20 DEC=20
MACRO1 MJ#(0) ARGF2
ARCON
MOVL C00189 V=8.0 ACC=20 DEC=20
MOVL C00190 V=8.0 ACC=20 DEC=20
MOVL C00191 V=8.0 ACC=20 DEC=20
MOVL C00192 V=8.0 ACC=20 DEC=20
MOVL C00193 V=8.0 ACC=20 DEC=20
MOVL C00194 V=8.0 ACC=20 DEC=20
MOVL C00195 V=8.0 ACC=20 DEC=20
MOVL C00196 V=8.0 ACC=20 DEC=20
MOVL C00197 V=8.0 ACC=20 DEC=20
MOVL C00198 V=8.0 ACC=20 DEC=20
MOVL C00199 V=8.0 ACC=20 DEC=20
MOVL C00200 V=8.0 ACC=20 DEC=20
MOVL C00201 V=8.0 ACC=20 DEC=20
MOVL C00202 V=8.0 ACC=20 DEC=20
MOVL C00203 V=8.0 ACC=20 DEC=20
MOVL C00204 V=8.0 ACC=20 DEC=20
MOVL C00205 V=8.0 ACC=20 DEC=20
MOVL C00206 V=8.0 ACC=20 DEC=20
MOVL C00207 V=8.0 ACC=20 DEC=20
MOVL C00208 V=8.0 ACC=20 DEC=20
MOVL C00209 V=8.0 ACC=20 DEC=20
MOVL C00210 V=8.0 ACC=20 DEC=20
MOVL C00211 V=8.0 ACC=20 DEC=20
MOVL C00212 V=8.0 ACC=20 DEC=20
MOVL C00213 V=8.0 ACC=20 DEC=20
MOVL C00214 V=8.0 ACC=20 DEC=20
MOVL C00215 V=8.0 ACC=20 DEC=20
MOVL C00216 V=8.0 ACC=20 DEC=20
MOVL C00217 V=8.0 ACC=20 DEC=20
MOVL C00218 V=8.0 ACC=20 DEC=20
ARCOF
TIMER T=60.0
MOVL C00219 V=11.0 ACC=20 DEC=20
MACRO1 MJ#(0) ARGF2
ARCON
MOVL C00220 V=8.0 ACC=20 DEC=20
MOVL C00221 V=8.0 ACC=20 DEC=20
MOVL C00222 V=8.0 ACC=20 DEC=20
MOVL C00223 V=8.0 ACC=20 DEC=20
MOVL C00224 V=8.0 ACC=20 DEC=20
MOVL C00225 V=8.0 ACC=20 DEC=20
MOVL C00226 V=8.0 ACC=20 DEC=20
MOVL C00227 V=8.0 ACC=20 DEC=20
MOVL C00228 V=8.0 ACC=20 DEC=20
MOVL C00229 V=8.0 ACC=20 DEC=20
MOVL C00230 V=8.0 ACC=20 DEC=20
MOVL C00231 V=8.0 ACC=20 DEC=20
MOVL C00232 V=8.0 ACC=20 DEC=20
MOVL C00233 V=8.0 ACC=20 DEC=20
MOVL C00234 V=8.0 ACC=20 DEC=20
MOVL C00235 V=8.0 ACC=20 DEC=20
MOVL C00236 V=8.0 ACC=20 DEC=20
MOVL C00237 V=8.0 ACC=20 DEC=20
MOVL C00238 V=8.0 ACC=20 DEC=20
MOVL C00239 V=8.0 ACC=20 DEC=20
MOVL C00240 V=8.0 ACC=20 DEC=20
MOVL C00241 V=8.0 ACC=20 DEC=20
MOVL C00242 V=8.0 ACC=20 DEC=20
MOVL C00243 V=8.0 ACC=20 DEC=20
MOVL C00244 V=8.0 ACC=20 DEC=20
MOVL C00245 V=8.0 ACC=20 DEC=20
MOVL C00246 V=8.0 ACC=20 DEC=20
MOVL C00247 V=8.0 ACC=20 DEC=20
MOVL C00248 V=8.0 ACC=20 DEC=20
MOVL C00249 V=8.0 ACC=20 DEC=20
ARCOF
TIMER T=60.0
MOVL C00250 V=11.0 ACC=20 DEC=20
MACRO1 MJ#(0) ARGF2
ARCON
MOVL C00251 V=8.0 ACC=20 DEC=20
MOVL C00252 V=8.0 ACC=20 DEC=20
MOVL C00253 V=8.0 ACC=20 DEC=20
MOVL C00254 V=8.0 ACC=20 DEC=20
MOVL C00255 V=8.0 ACC=20 DEC=20
MOVL C00256 V=8.0 ACC=20 DEC=20
MOVL C00257 V=8.0 ACC=20 DEC=20
MOVL C00258 V=8.0 ACC=20 DEC=20
MOVL C00259 V=8.0 ACC=20 DEC=20
MOVL C00260 V=8.0 ACC=20 DEC=20
MOVL C00261 V=8.0 ACC=20 DEC=20
MOVL C00262 V=8.0 ACC=20 DEC=20
MOVL C00263 V=8.0 ACC=20 DEC=20
MOVL C00264 V=8.0 ACC=20 DEC=20
MOVL C00265 V=8.0 ACC=20 DEC=20
MOVL C00266 V=8.0 ACC=20 DEC=20
MOVL C00267 V=8.0 ACC=20 DEC=20
MOVL C00268 V=8.0 ACC=20 DEC=20
MOVL C00269 V=8.0 ACC=20 DEC=20
MOVL C00270 V=8.0 ACC=20 DEC=20
MOVL C00271 V=8.0 ACC=20 DEC=20
MOVL C00272 V=8.0 ACC=20 DEC=20
MOVL C00273 V=8.0 ACC=20 DEC=20
MOVL C00274 V=8.0 ACC=20 DEC=20
MOVL C00275 V=8.0 ACC=20 DEC=20
MOVL C00276 V=8.0 ACC=20 DEC=20
MOVL C00277 V=8.0 ACC=20 DEC=20
MOVL C00278 V=8.0 ACC=20 DEC=20
MOVL C00279 V=8.0 ACC=20 DEC=20
MOVL C00280 V=8.0 ACC=20 DEC=20
ARCOF
TIMER T=60.0
MOVL C00281 V=11.0 ACC=20 DEC=20
MACRO1 MJ#(0) ARGF2
ARCON
MOVL C00282 V=8.0 ACC=20 DEC=20
MOVL C00283 V=8.0 ACC=20 DEC=20
MOVL C00284 V=8.0 ACC=20 DEC=20
MOVL C00285 V=8.0 ACC=20 DEC=20
MOVL C00286 V=8.0 ACC=20 DEC=20
MOVL C00287 V=8.0 ACC=20 DEC=20
MOVL C00288 V=8.0 ACC=20 DEC=20
MOVL C00289 V=8.0 ACC=20 DEC=20
MOVL C00290 V=8.0 ACC=20 DEC=20
MOVL C00291 V=8.0 ACC=20 DEC=20
MOVL C00292 V=8.0 ACC=20 DEC=20
MOVL C00293 V=8.0 ACC=20 DEC=20
MOVL C00294 V=8.0 ACC=20 DEC=20
MOVL C00295 V=8.0 ACC=20 DEC=20
MOVL C00296 V=8.0 ACC=20 DEC=20
MOVL C00297 V=8.0 ACC=20 DEC=20
MOVL C00298 V=8.0 ACC=20 DEC=20
MOVL C00299 V=8.0 ACC=20 DEC=20
MOVL C00300 V=8.0 ACC=20 DEC=20
MOVL C00301 V=8.0 ACC=20 DEC=20
MOVL C00302 V=8.0 ACC=20 DEC=20
MOVL C00303 V=8.0 ACC=20 DEC=20
MOVL C00304 V=8.0 ACC=20 DEC=20
MOVL C00305 V=8.0 ACC=20 DEC=20
MOVL C00306 V=8.0 ACC=20 DEC=20
MOVL C00307 V=8.0 ACC=20 DEC=20
MOVL C00308 V=8.0 ACC=20 DEC=20
MOVL C00309 V=8.0 ACC=20 DEC=20
MOVL C00310 V=8.0 ACC=20 DEC=20
MOVL C00311 V=8.0 ACC=20 DEC=20
ARCOF
TIMER T=60.0
MOVL C00312 V=11.0 ACC=20 DEC=20
MACRO1 MJ#(0) ARGF2
ARCON
MOVL C00313 V=8.0 ACC=20 DEC=20
MOVL C00314 V=8.0 ACC=20 DEC=20
MOVL C00315 V=8.0 ACC=20 DEC=20
MOVL C00316 V=8.0 ACC=20 DEC=20
MOVL C00317 V=8.0 ACC=20 DEC=20
MOVL C00318 V=8.0 ACC=20 DEC=20
MOVL C00319 V=8.0 ACC=20 DEC=20
MOVL C00320 V=8.0 ACC=20 DEC=20
MOVL C00321 V=8.0 ACC=20 DEC=20
MOVL C00322 V=8.0 ACC=20 DEC=20
MOVL C00323 V=8.0 ACC=20 DEC=20
MOVL C00324 V=8.0 ACC=20 DEC=20
MOVL C00325 V=8.0 ACC=20 DEC=20
MOVL C00326 V=8.0 ACC=20 DEC=20
MOVL C00327 V=8.0 ACC=20 DEC=20
MOVL C00328 V=8.0 ACC=20 DEC=20
MOVL C00329 V=8.0 ACC=20 DEC=20
MOVL C00330 V=8.0 ACC=20 DEC=20
MOVL C00331 V=8.0 ACC=20 DEC=20
MOVL C00332 V=8.0 ACC=20 DEC=20
MOVL C00333 V=8.0 ACC=20 DEC=20
MOVL C00334 V=8.0 ACC=20 DEC=20
MOVL C00335 V=8.0 ACC=20 DEC=20
MOVL C00336 V=8.0 ACC=20 DEC=20
MOVL C00337 V=8.0 ACC=20 DEC=20
MOVL C00338 V=8.0 ACC=20 DEC=20
MOVL C00339 V=8.0 ACC=20 DEC=20
MOVL C00340 V=8.0 ACC=20 DEC=20
MOVL C00341 V=8.0 ACC=20 DEC=20
MOVL C00342 V=8.0 ACC=20 DEC=20
ARCOF
TIMER T=60.0
MOVL C00343 V=11.0 ACC=20 DEC=20
MACRO1 MJ#(0) ARGF2
ARCON
MOVL C00344 V=8.0 ACC=20 DEC=20
MOVL C00345 V=8.0 ACC=20 DEC=20
MOVL C00346 V=8.0 ACC=20 DEC=20
MOVL C00347 V=8.0 ACC=20 DEC=20
MOVL C00348 V=8.0 ACC=20 DEC=20
MOVL C00349 V=8.0 ACC=20 DEC=20
MOVL C00350 V=8.0 ACC=20 DEC=20
MOVL C00351 V=8.0 ACC=20 DEC=20
MOVL C00352 V=8.0 ACC=20 DEC=20
MOVL C00353 V=8.0 ACC=20 DEC=20
MOVL C00354 V=8.0 ACC=20 DEC=20
MOVL C00355 V=8.0 ACC=20 DEC=20
MOVL C00356 V=8.0 ACC=20 DEC=20
MOVL C00357 V=8.0 ACC=20 DEC=20
MOVL C00358 V=8.0 ACC=20 DEC=20
MOVL C00359 V=8.0 ACC=20 DEC=20
MOVL C00360 V=8.0 ACC=20 DEC=20
MOVL C00361 V=8.0 ACC=20 DEC=20
MOVL C00362 V=8.0 ACC=20 DEC=20
MOVL C00363 V=8.0 ACC=20 DEC=20
MOVL C00364 V=8.0 ACC=20 DEC=20
MOVL C00365 V=8.0 ACC=20 DEC=20
MOVL C00366 V=8.0 ACC=20 DEC=20
MOVL C00367 V=8.0 ACC=20 DEC=20
MOVL C00368 V=8.0 ACC=20 DEC=20
MOVL C00369 V=8.0 ACC=20 DEC=20
MOVL C00370 V=8.0 ACC=20 DEC=20
MOVL C00371 V=8.0 ACC=20 DEC=20
MOVL C00372 V=8.0 ACC=20 DEC=20
MOVL C00373 V=8.0 ACC=20 DEC=20
ARCOF
TIMER T=60.0
MOVL C00374 V=11.0 ACC=20 DEC=20
MACRO1 MJ#(0) ARGF2
ARCON
MOVL C00375 V=8.0 ACC=20 DEC=20
MOVL C00376 V=8.0 ACC=20 DEC=20
MOVL C00377 V=8.0 ACC=20 DEC=20
MOVL C00378 V=8.0 ACC=20 DEC=20
MOVL C00379 V=8.0 ACC=20 DEC=20
MOVL C00380 V=8.0 ACC=20 DEC=20
MOVL C00381 V=8.0 ACC=20 DEC=20
MOVL C00382 V=8.0 ACC=20 DEC=20
MOVL C00383 V=8.0 ACC=20 DEC=20
MOVL C00384 V=8.0 ACC=20 DEC=20
MOVL C00385 V=8.0 ACC=20 DEC=20
MOVL C00386 V=8.0 ACC=20 DEC=20
MOVL C00387 V=8.0 ACC=20 DEC=20
MOVL C00388 V=8.0 ACC=20 DEC=20
MOVL C00389 V=8.0 ACC=20 DEC=20
MOVL C00390 V=8.0 ACC=20 DEC=20
MOVL C00391 V=8.0 ACC=20 DEC=20
MOVL C00392 V=8.0 ACC=20 DEC=20
MOVL C00393 V=8.0 ACC=20 DEC=20
MOVL C00394 V=8.0 ACC=20 DEC=20
MOVL C00395 V=8.0 ACC=20 DEC=20
MOVL C00396 V=8.0 ACC=20 DEC=20
MOVL C00397 V=8.0 ACC=20 DEC=20
MOVL C00398 V=8.0 ACC=20 DEC=20
MOVL C00399 V=8.0 ACC=20 DEC=20
MOVL C00400 V=8.0 ACC=20 DEC=20
MOVL C00401 V=8.0 ACC=20 DEC=20
MOVL C00402 V=8.0 ACC=20 DEC=20
MOVL C00403 V=8.0 ACC=20 DEC=20
MOVL C00404 V=8.0 ACC=20 DEC=20
ARCOF
TIMER T=60.0
MOVL C00405 V=11.0 ACC=20 DEC=20
MACRO1 MJ#(0) ARGF2
ARCON
MOVL C00406 V=8.0 ACC=20 DEC=20
MOVL C00407 V=8.0 ACC=20 DEC=20
MOVL C00408 V=8.0 ACC=20 DEC=20
MOVL C00409 V=8.0 ACC=20 DEC=20
MOVL C00410 V=8.0 ACC=20 DEC=20
MOVL C00411 V=8.0 ACC=20 DEC=20
MOVL C00412 V=8.0 ACC=20 DEC=20
MOVL C00413 V=8.0 ACC=20 DEC=20
MOVL C00414 V=8.0 ACC=20 DEC=20
MOVL C00415 V=8.0 ACC=20 DEC=20
MOVL C00416 V=8.0 ACC=20 DEC=20
MOVL C00417 V=8.0 ACC=20 DEC=20
MOVL C00418 V=8.0 ACC=20 DEC=20
MOVL C00419 V=8.0 ACC=20 DEC=20
MOVL C00420 V=8.0 ACC=20 DEC=20
MOVL C00421 V=8.0 ACC=20 DEC=20
MOVL C00422 V=8.0 ACC=20 DEC=20
MOVL C00423 V=8.0 ACC=20 DEC=20
MOVL C00424 V=8.0 ACC=20 DEC=20
MOVL C00425 V=8.0 ACC=20 DEC=20
MOVL C00426 V=8.0 ACC=20 DEC=20
MOVL C00427 V=8.0 ACC=20 DEC=20
MOVL C00428 V=8.0 ACC=20 DEC=20
MOVL C00429 V=8.0 ACC=20 DEC=20
MOVL C00430 V=8.0 ACC=20 DEC=20
MOVL C00431 V=8.0 ACC=20 DEC=20
MOVL C00432 V=8.0 ACC=20 DEC=20
MOVL C00433 V=8.0 ACC=20 DEC=20
MOVL C00434 V=8.0 ACC=20 DEC=20
MOVL C00435 V=8.0 ACC=20 DEC=20
ARCOF
TIMER T=60.0
MOVL C00436 V=11.0 ACC=20 DEC=20
MOVJ C00437 VJ=0.78
END
